(* Logix 5000 project; controller lab5BnB 5069-L306ERM rev 38.11; software revision 38.02 *)

TASK MainTask (periodic, rate 1 ms, priority 10, watchdog 1 ms) : MainProgram

MODULES
   Local : 5069-L306ERM (5069 0, rev 38.11)
       : 5069-OB16 (5069 2, rev 3.13, StandardDataDriven RPI 5 ms)
       : 5069-IB16 (5069 1, rev 2.16, StandardDataDriven RPI 5 ms)
       : vendor 1 type 115 code 320 (5069 4, rev 2.13, StandardDataDriven RPI 1 ms)
       : 5069-IF8 (5069 3, rev 3.11, StandardDataDriven RPI 1 ms)
END_MODULES

ADD_ON_INSTRUCTION Angle_Controller   (* revision 1.0 *)
VAR_INPUT
   Kp : REAL; {access None}
   Kd : REAL; {access None}
   Ki : REAL; {access None}
END_VAR
VAR_OUTPUT
   MotorInInt : REAL; {access None}
END_VAR
VAR_INPUT
   MotorVoltageInt : REAL; {access None}
   DesiredMotorAngleDeg : REAL; {access None}
END_VAR
VAR
   DERV_01 : DERIVATIVE;
   INTG_02 : INTEGRATOR;
   LPF_01 : FILTER_LOW_PASS;
   MUL_01 : FBD_MATH;
   SCL_01 : SCALE;
   SCL_02 : SCALE;
   SSUM_01 : SELECTED_SUMMER;
   SUB_01 : FBD_MATH;
   BalanceMax : REAL; {access None}
   BalanceMin : REAL; {access None}
   MotorAngleDeg : REAL; {access None}
   MyError : REAL; {access None}
   PreFilter : REAL; {access None}
   PostFilter : REAL; {access None}
   __lECF02074BD2460E6 : REAL; {access None}
   __l28C6010D865A5A33 : REAL; {access None}
   __l0884565386038A91 : REAL; {access None}
   __l2DF07EE77D244EFB : REAL; {access None}
   __l1766871E0CB1B884 : REAL; {access None}
   __l0E750273472B5D8B : REAL; {access None}
   __lD887463BECBAFEBD : REAL; {access None}
   __l08A3F56F66BAD335 : REAL; {access None}
END_VAR

ROUTINE Logic   (* function block diagram *)
   SHEET 1
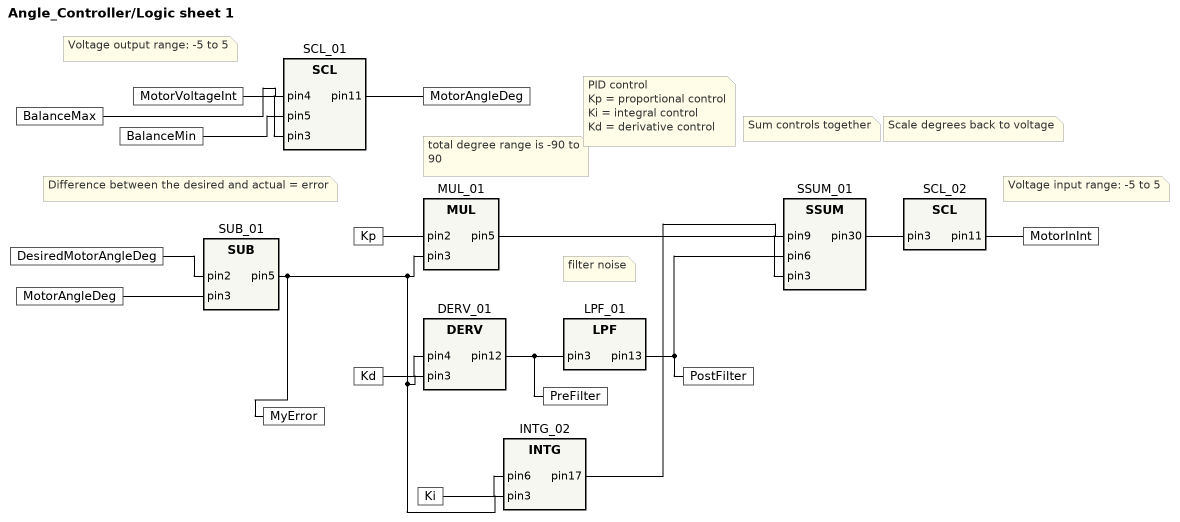
   // Difference between the desired and actual = error
   // Voltage output range: -5 to 5
   // total degree range is -90 to
   // 90
   // filter noise
   // PID control
   // Kp = proportional control
   // Ki = integral control
   // Kd = derivative control
   // Sum controls together
   // Scale degrees back to voltage
   // Voltage input range: -5 to 5
   SUB_01 : SUB(pin2 := DesiredMotorAngleDeg, pin3 := MotorAngleDeg);
   MyError := SUB_01.pin5;
   SCL_01 : SCL(pin3 := MotorVoltageInt, pin4 := BalanceMax, pin5 := BalanceMin);
   MotorAngleDeg := SCL_01.pin11;
   MUL_01 : MUL(pin2 := Kp, pin3 := SUB_01.pin5);
   DERV_01 : DERV(pin3 := SUB_01.pin5, pin4 := Kd);
   INTG_02 : INTG(pin3 := SUB_01.pin5, pin6 := Ki);
   PreFilter := DERV_01.pin12;
   LPF_01 : LPF(pin3 := DERV_01.pin12);
   PostFilter := LPF_01.pin13;
   SSUM_01 : SSUM(pin3 := MUL_01.pin5, pin6 := LPF_01.pin13, pin9 := INTG_02.pin17);
   SCL_02 : SCL(pin3 := SSUM_01.pin30);
   MotorInInt := SCL_02.pin11;
END_ROUTINE
END_ADD_ON_INSTRUCTION

ADD_ON_INSTRUCTION Position_Controller   (* revision 1.0 *)
VAR_INPUT
   Kp_position : REAL; {visible}
   Kd_position : REAL; {visible}
   Ki_position : REAL; {visible}
   Actual_Position : REAL; {visible}
   Desired_Position : REAL; {visible}
END_VAR
VAR_OUTPUT
   angle_out : REAL; {visible}
END_VAR
VAR
   SCL_01 : SCALE; {access None}
   Desired_Position_Inches : DINT; {access None}
   SCL_02 : SCALE; {access None}
   Actual_Position_Inches : DINT; {access None}
   SUB_01 : FBD_MATH;
   MyErrorPosition : DINT; {access None}
   MUL_01 : FBD_MATH;
   SCL_03 : SCALE;
   DERV_01 : DERIVATIVE; {access None}
   INTG_01 : INTEGRATOR; {access None}
   SSUM_01 : SELECTED_SUMMER; {access None}
   LPF_02 : FILTER_LOW_PASS; {access None}
   LPF_03 : FILTER_LOW_PASS; {access None}
   __l331A2C5B709CA8A7 : REAL; {access None}
   __l8C615611B29A5C42 : REAL; {access None}
   __l35E6236049371C91 : REAL; {access None}
   __l45EB0282393F6911 : REAL; {access None}
   __l367F46D6FCA640C7 : REAL; {access None}
END_VAR

ROUTINE Logic   (* function block diagram *)
   SHEET 1
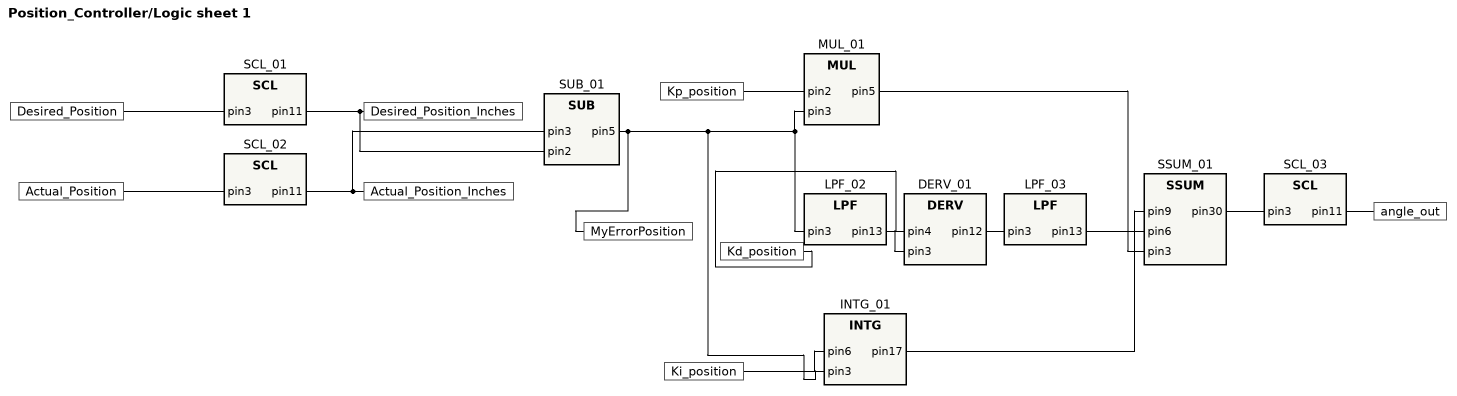
   SCL_01 : SCL(pin3 := Desired_Position);
   SCL_02 : SCL(pin3 := Actual_Position);
   Desired_Position_Inches := SCL_01.pin11;
   Actual_Position_Inches := SCL_02.pin11;
   SUB_01 : SUB(pin2 := SCL_01.pin11, pin3 := SCL_02.pin11);
   MyErrorPosition := SUB_01.pin5;
   MUL_01 : MUL(pin2 := Kp_position, pin3 := SUB_01.pin5);
   LPF_02 : LPF(pin3 := SUB_01.pin5);
   INTG_01 : INTG(pin3 := SUB_01.pin5, pin6 := Ki_position);
   DERV_01 : DERV(pin3 := LPF_02.pin13, pin4 := Kd_position);
   LPF_03 : LPF(pin3 := DERV_01.pin12);
   SSUM_01 : SSUM(pin3 := MUL_01.pin5, pin6 := LPF_03.pin13, pin9 := INTG_01.pin17);
   SCL_03 : SCL(pin3 := SSUM_01.pin30);
   angle_out := SCL_03.pin11;
END_ROUTINE
END_ADD_ON_INSTRUCTION

VAR_GLOBAL   (* controller tags *)
   DesiredMotorAngleDeg : REAL := 4.358898;
   DesiredPosition : ALIAS FOR Local:3:I.Ch02.Data;
   DesiredPositionInches : REAL := -2.6956902;
   Kd : REAL := 0.8;
   Kd_Position : REAL := 8.0;
   Ki : REAL := 0.5;
   Ki_Position : REAL := 10.0;
   Kp : REAL := 0.4;
   Kp_Position : REAL := 10.0;
   MotorAngleDeg : REAL := 0.4554901;
   MotorInInt : ALIAS FOR Local:4:O.Ch00.Data;
   MotorVoltageInt : ALIAS FOR Local:3:I.Ch00.Data;
   Position : ALIAS FOR Local:3:I.Ch01.Data;
   PositionInches : REAL := -2.6805582;
END_VAR

PROGRAM MainProgram   (* main routine main *)
VAR
   Angle_Controller_01 : Angle_Controller;
   Position_Controller_01 : Position_Controller;
   SCL_01 : SCALE;
   SCL_02 : SCALE; {access None}
   SCL_03 : SCALE; {access None}
END_VAR

ROUTINE main   (* function block diagram *)
   SHEET 1
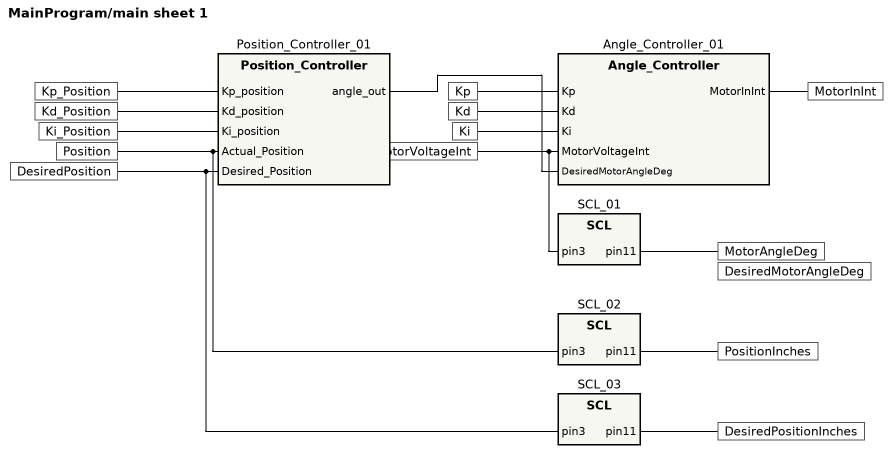
   Position_Controller_01 : Position_Controller(Kp_position := Kp_Position, Kd_position := Kd_Position, Ki_position := Ki_Position, Actual_Position := Position, Desired_Position := DesiredPosition);
   Angle_Controller_01 : Angle_Controller(Kp := Kp, Kd := Kd, Ki := Ki, MotorVoltageInt := MotorVoltageInt, DesiredMotorAngleDeg := Position_Controller_01.angle_out);
   SCL_01 : SCL(pin3 := MotorVoltageInt);
   SCL_02 : SCL(pin3 := Position);
   SCL_03 : SCL(pin3 := DesiredPosition);
   MotorAngleDeg := SCL_01.pin11;
   // unwired output reference DesiredMotorAngleDeg
   PositionInches := SCL_02.pin11;
   DesiredPositionInches := SCL_03.pin11;
   MotorInInt := Angle_Controller_01.MotorInInt;
END_ROUTINE
END_PROGRAM
